Fanuc KAREL source: kb00051.KL

PROGRAM KB00051
%STACKSIZE=65535
%PRIORITY=65535
%NOLOCKGROUP
VAR
P1 : INTEGER
P2 : INTEGER
RESULT : JOINTPOS9
BEGIN
P1=1
P2=1
-- UNRESOLVED_PC line 10 opcodes [27 22 22 27 9D 76 7E 4A] marker_code=24
END KB00051
